TYPE E_MqttObservedHaStatus :
(
    Unknown,
    Offline,
    Online
);
END_TYPE

(* stored: Version 1.1.0.1
   DUT E_MqttObservedHaStatus: Id {4c0c3919-b7ec-41a6-bdd7-039d14fc0ba5} *)
